TYPE "DT_DIGITAL_OUTPUTS_ALL"
VERSION : 0.1
   STRUCT
      TUR_FRA_KAP_CROSS : "DT_DIGITAL_OUTPUT_TUR_FRANCIS_KAPLAN_CROSS";
      TUR_PELT_DEFLECT : "DT_DIGITAL_OUTPUT_TUR_PELTON_DEFLECTOR";
      TUR_PELT_NOZZLE : "DT_DIGITAL_OUTPUT_TUR_PELTON_NOZZLE";
      TUR_OTHER : "DT_DIGITAL_OUTPUT_TUR_OTHER";
      SUBSYS : "DT_DIGITAL_OUTPUT_SUBSYSTEMS";
      CTRL_SYNC_EXC : "DT_DIGITAL_OUTPUT_CTRL_SYNC_EXC";
      WATERWAY_INTAKE : "DT_DIGITAL_OUTPUT_WATERWAY_AND_INTAKE";
      CUBIC_AND_SIGNAL : "DT_DIGITAL_OUTPUT_CUBICLES_AND_SIGNALIZATION";
      SN : "DT_DIGITAL_OUTPUT_SN";
   END_STRUCT;

END_TYPE

